(* IEC 61131-3 sources: SRCI_CLIENT_PLC/RobotLibrary/Library/POUs/Trigger/MC_SetTriggerRegister/Structures, 4 files *)

(* ---- SetTriggerRegisterOutCmd.st ---- *)
{attribute 'pack_mode' := '1'}
// -------------------------------------------------------------------------
//  SRCI Robot Library
// -------------------------------------------------------------------------
//
//  Object:      SetTriggerRegisterOutCmd
//  Author:      Thorsten Brach
//  Date:        2024-08-03
//
//  Description:
//
//
//  Copyright:
//    (C) 2024 Thorsten Brach. All rights reserved
//             Licensed under the MIT License.
//
//  Disclaimer:
//    This project is provided without any guarantee and can be used for
//    private and commercial purposes. Any use is at the user’s
//    own risk and responsibility.
//
// -------------------------------------------------------------------------
TYPE SetTriggerRegisterOutCmd :
STRUCT
  /// Unique system-generated ID of the "Action" when the function is triggered.
  /// • >0: The "Action" is started by the trigger function with identical FollowID.
  /// • <0: The "Action" is stopped by the trigger function with identical FollowID.
  /// For more information see chapter 5.5.12.4 EmitterID, ListenerID, FollowID and OriginID
  OriginID               : INT;
  /// Relates to ListenerID >0
  /// Number of successful trigger -based command invocations
  /// For more information refer to chapter 5.5.12.4.
  InvocationCounter      : USINT;
  /// Unique system-generated ID of the trigger function when the function is called by user.
  /// For more information see chapter 5.5.12.4.
  FollowID               : DINT;
END_STRUCT
END_TYPE

(* ---- SetTriggerRegisterParCmd.st ---- *)
{attribute 'pack_mode' := '1'}
// -------------------------------------------------------------------------
//  SRCI Robot Library
// -------------------------------------------------------------------------
//
//  Object:      SetTriggerRegisterParCmd
//  Author:      Thorsten Brach
//  Date:        2024-08-03
//
//  Description:
//
//
//  Copyright:
//    (C) 2024 Thorsten Brach. All rights reserved
//             Licensed under the MIT License.
//
//  Disclaimer:
//    This project is provided without any guarantee and can be used for
//    private and commercial purposes. Any use is at the user’s
//    own risk and responsibility.
//
// -------------------------------------------------------------------------
TYPE SetTriggerRegisterParCmd :
STRUCT
  /// Specifies the trigger event according to Table 6-596.
  /// For more information about registers on the RC see chapters 6.4.4 and 6.4.5.
  TriggerMode            : TriggerModeIo;
  /// Determines whether the start condition is evaluated or not.
  /// • FALSE: Start condition is not evaluated (default).
  /// • TRUE: Start condition is evaluated.
  EvaluateStartCondition : BOOL;
  /// Depending on "TriggerMode":
  /// • Digital (refers to "TriggerMode" 10-13, 20-23): Specifies the desired byte address of the input or output signal that shall be read.
  /// • Analog/Integer/Real (refers to "TriggerMode" 30-37, 40-47, 50-57, 60- 67): Specifies the target values that shall be read.
  /// For more information about registers refer to Figure 6-206.
  Index                  : USINT;
  /// Depending on "TriggerMode":
  /// • Digital (refers to TriggerMode 10-13,20-23): Specifies the desired bit address of the input or output signal that shall be read.
  /// • Analog/Integer/Real (refers to TriggerMode 30-37, 40-47, 50-57, 60- 67): Not relevant and deactivated for user input.
  /// For more information about registers refer to Figure 6-206
  BitIndex               : USINT;
  /// Reference integer value, for triggering the Action function with the EmitterID.
  /// • Relates to "TriggerMode" 50-57
  IntValue               : ARRAY[1..2] OF INT;
  /// Reference real value, analog input or output value, for triggering the Action function with the EmitterID.
  /// • Relates to "TriggerMode" 30-37, 40-47,60-67
  RealValue              : ARRAY[1..2] OF REAL;
  /// ID of associated trigger function:
  /// • 0: Immediately (default). - Start executing this function immediately.
  /// • >0: Trigger - Start executing, when the trigger function with the identical EmitterID is triggered.
  /// Always positive.
  /// For more information, see chapter 5.5.12 Triggers
  ListenerID             : SINT;
  /// ID of the Action function that will be executed when the trigger condition is met
  /// • >0: Start Action        - Start executing the Action function with the identical ListenerID.
  /// • <0: Stop Action         - Stop executing the Action function with the identical ListenerID.
  /// •  0: Undefined (default) - If no EmitterID is defined, the function returns an error message
  /// For more information see chapter 5.5.12.4
  EmitterID              : SINT;
END_STRUCT
END_TYPE

(* ---- SetTriggerRegisterRecvData.st ---- *)
{attribute 'pack_mode' := '1'}
// -------------------------------------------------------------------------
//  SRCI Robot Library
// -------------------------------------------------------------------------
//
//  Object:      SetTriggerRegisterRecvData
//  Author:      Thorsten Brach
//  Date:        2024-08-03
//
//  Description:
//
//
//  Copyright:
//    (C) 2024 Thorsten Brach. All rights reserved
//             Licensed under the MIT License.
//
//  Disclaimer:
//    This project is provided without any guarantee and can be used for
//    private and commercial purposes. Any use is at the user’s
//    own risk and responsibility.
//
// -------------------------------------------------------------------------
TYPE SetTriggerRegisterRecvData EXTENDS RspHeader :
STRUCT
  /// Relates to ListenerID >0
  /// Number of successful trigger -based command invocations
  /// For more information refer to chapter 5.5.12.4.
  InvocationCounter      : USINT;
  /// Reserve
  Reserve                : SINT;
  /// Unique system-generated ID of the "Action" when the function is triggered.
  /// • >0: The "Action" is started by the trigger function with identical FollowID.
  /// • <0: The "Action" is stopped by the trigger function with identical FollowID.
  /// For more information see chapter 5.5.12.4 EmitterID, ListenerID, FollowID and OriginID
  OriginID               : INT;
END_STRUCT
END_TYPE

(* ---- SetTriggerRegisterSendData.st ---- *)
{attribute 'pack_mode' := '1'}
// -------------------------------------------------------------------------
//  SRCI Robot Library
// -------------------------------------------------------------------------
//
//  Object:      SetTriggerRegisterSendData
//  Author:      Thorsten Brach
//  Date:        2024-08-03
//
//  Description:
//
//
//  Copyright:
//    (C) 2024 Thorsten Brach. All rights reserved
//             Licensed under the MIT License.
//
//  Disclaimer:
//    This project is provided without any guarantee and can be used for
//    private and commercial purposes. Any use is at the user’s
//    own risk and responsibility.
//
// -------------------------------------------------------------------------
TYPE SetTriggerRegisterSendData EXTENDS CmdHeader:
STRUCT
  /// ID of Action that will be executed when this command is active
  /// • >0: Start Action - Start executing the Action function with the identical ListenerID.
  /// • <0: Stop Action  -  Stop executing the Action function with the identical ListenerID.
  /// • 0: No trigger (default)-  If no EmitterID is defined, the function will not trigger any Action during its execution
  /// For more information see section Triggers of this chapter or chapter 5.5.12.4.
  EmitterID              : ARRAY [0..3] OF SINT;
  /// ID of associated trigger function:
  /// • 0: Immediately (default) - Start executing this function immediately.
  /// • >0: Trigger -  Start executing, when the trigger function with the identical EmitterID is triggered.
  /// Always positive.
  /// For more information, see chapter 5.5.12 Triggers
  ListenerID             : SINT;
  /// Reserve
  Reserve                : SINT;
  /// Reference integer value, for triggering the Action function with the EmitterID.
  /// • Relates to "TriggerMode" 50-57
  IntValue               : ARRAY[1..2] OF INT;
  /// Reference real value, analog input or output value, for triggering the Action function with the EmitterID.
  /// • Relates to "TriggerMode" 30-37, 40-47,60-67
  RealValue              : ARRAY[1..2] OF REAL;
  /// Specifies the trigger event according to Table 6-596.
  /// For more information about registers on the RC see chapters 6.4.4 and 6.4.5.
  TriggerMode            : SINT;
  /// Depending on "TriggerMode":
  /// • Digital (refers to "TriggerMode" 10-13, 20-23): Specifies the desired byte address of the input or output signal that shall be read.
  /// • Analog/Integer/Real (refers to "TriggerMode" 30-37, 40-47, 50-57, 60- 67): Specifies the target values that shall be read.
  /// For more information about registers refer to Figure 6-206.
  Index                  : USINT;
  /// Depending on "TriggerMode":
  /// • Digital (refers to TriggerMode 10-13,20-23): Specifies the desired bit address of the input or output signal that shall be read.
  /// • Analog/Integer/Real (refers to TriggerMode 30-37, 40-47, 50-57, 60- 67): Not relevant and deactivated for user input.
  /// For more information about registers refer to Figure 6-206
  BitIndex               : USINT;
END_STRUCT
END_TYPE
